// SIMATIC S7-200 project (STEP 7-Micro/WIN), CPU 224 CN REL 02.01

SYMBOL_TABLE ????1
boton_sb1        I1.3
boton_sb2        I1.2
selector         I1.5
parada           I1.4
act1             Q0.0
act2             Q0.2
act3             Q0.3
act4             ?0_40_0
END_SYMBOL_TABLE

ORGANIZATION_BLOCK ???:OB1
TITLE=????
BEGIN
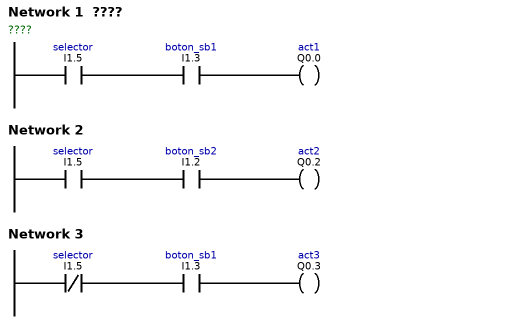
Network 1 // ????
// ????
LD     selector:I1.5
A      boton_sb1:I1.3
=      act1:Q0.0
Network 2
LD     selector:I1.5
A      boton_sb2:I1.2
=      act2:Q0.2
Network 3
LDN    selector:I1.5
A      boton_sb1:I1.3
=      act3:Q0.3
END_ORGANIZATION_BLOCK
